// ---- Machine/FB_Centering.TcPOU
// Centraggio TL/TB di Aut260045 (ex passi 55-78 di MAIN.StateMachine, stessi numeri in nStep).
// Corsa rapida IN STROKE, ricerca dei pezzi fino a MAX STROKE con chiusura dei palpatori, arresto,
// chiusura morsa e corsa EXTRA, risalita dei centratori. Usa direttamente I/O e parametri del programma:
// e' un modulo della macchina, non del Core.
// Va chiamato a ogni ciclo PLC (gli FB di movimento e i timer devono girare sempre); con bExecute
// esegue, senza torna a Idle. Gli allarmi li memorizza qui (RaiseAlarm); il ciclo legge bDone, bFailed, bAbort.
FUNCTION_BLOCK FB_Centering
VAR_INPUT
	bExecute		: BOOL;				// il ciclo e' nel passo Centering
	bStart			: BOOL;				// consenso start (attese del passo-passo)
	bStepMode		: BOOL;				// passo-passo: tra le fasi si aspetta lo start
	fMoveSpeed		: LREAL := 200;		// velocita' USE nelle corse IN STROKE ed EXTRA
	fSearchSpeed	: LREAL := 30;		// velocita' USE nella ricerca dei pezzi
	nGroupIdBase	: UDINT := 7;		// ID NC dei gruppi da svuotare prima delle corse PTP
END_VAR
VAR_IN_OUT
	stUseL			: AXIS_REF;
	stUseR			: AXIS_REF;
END_VAR
VAR_OUTPUT
	nStep			: E_CenteringStep;
	bDone			: BOOL;		// centraggio finito: fMeasureL/R valide
	bFailed			: BOOL;		// pezzo gia' presente o non trovato: si rifa' il posizionamento iniziale
	bAbort			: BOOL;		// errore NC: il ciclo va in abort
	fMeasureL		: LREAL;	// corsa di ricerca SX (inizio - fine), per la tolleranza TB
	fMeasureR		: LREAL;
END_VAR
VAR
	fbClearGroup	: ARRAY[0..2] OF CfgReconfigGroup;
	fbMoveL			: MC_MoveAbsolute;
	fbMoveR			: MC_MoveAbsolute;
	fbStopL			: MC_Halt;
	fbStopR			: MC_Halt;
	fbClampsDelay	: TON;
	fbTlClampsDelay	: TON;
	fbUpDownDelay	: TON;
	fStrokeInL		: LREAL;
	fStrokeInR		: LREAL;
	fStartL			: LREAL;
	fStartR			: LREAL;
	fMaxStrokeL		: LREAL;
	fMaxStrokeR		: LREAL;
	fEndL			: LREAL;
	fEndR			: LREAL;
	fExtraL			: LREAL;
	fExtraR			: LREAL;
	pz1Found		: BOOL;
	pz2Found		: BOOL;
	pz3Found		: BOOL;
	pz4Found		: BOOL;
	i				: UINT;
END_VAR

// Valori di riposo a ogni ciclo (prima in MAIN.InitCyclic): i passi li riaccendono.
fbStopL.Execute := FALSE;
fbStopR.Execute := FALSE;
fbMoveL.Execute := FALSE;
fbMoveL.Velocity := 0;
fbMoveR.Execute := FALSE;
fbMoveR.Velocity := 0;
fbClampsDelay.IN := FALSE;
fbClampsDelay.PT := T#800MS;
fbTlClampsDelay.IN := FALSE;
fbTlClampsDelay.PT := T#250MS;
fbUpDownDelay.IN := FALSE;
fbUpDownDelay.PT := T#800MS;
bDone := FALSE;
bFailed := FALSE;
bAbort := FALSE;

IF NOT bExecute THEN
	nStep := E_CenteringStep.Idle;
ELSIF nStep = E_CenteringStep.Idle THEN
	nStep := E_CenteringStep.ClearGroups;
END_IF

CASE nStep OF
	(******************* Clear groups for centering *******************)  
	E_CenteringStep.ClearGroups:
		FOR i:=0 TO 2 DO
			fbClearGroup[i](
				nGroupId:=nGroupIdBase+i,
				bExecute:=TRUE,
				tTimeOut:=T#100MS );
		END_FOR
		
		IF (NOT fbClearGroup[0].bBusy) AND (NOT fbClearGroup[1].bBusy) AND (NOT fbClearGroup[2].bBusy) THEN
			fbClearGroup[0]( bExecute:=FALSE );
			fbClearGroup[1]( bExecute:=FALSE );
			fbClearGroup[2]( bExecute:=FALSE );
			nStep := E_CenteringStep.ApproachPrepare;
			
			//IO.centeringLeft1Set := FALSE;
			//IO.centeringLeft2Set := FALSE;
			//IO.centeringLeft3Set := FALSE;
			//IO.centeringLeft4Set := FALSE;
			io.centeringOutSet := TRUE;
		END_IF
		
		IF fbClearGroup[0].bErr OR fbClearGroup[1].bErr OR fbClearGroup[2].bErr THEN
			RaiseAlarm(Id := E_Alarm.NcCenteringClearGroup, Info := MAX(fbClearGroup[0].nErrId, fbClearGroup[1].nErrId, fbClearGroup[2].nErrId));
			bAbort := TRUE;
			nStep := E_CenteringStep.Error;
		END_IF
	
	(*************** Prepare fast in stroke movement ***************)  
	E_CenteringStep.ApproachPrepare:	
		fStrokeInL := stUseL.NcToPlc.ActPos - ProgramDB.parameters.inStrokeL;
		fStrokeInR := stUseR.NcToPlc.ActPos - ProgramDB.parameters.inStrokeR;
	    fbMoveL(Axis := stUseL, Execute := FALSE);
		fbMoveR(Axis := stUseR, Execute := FALSE);
		nStep := E_CenteringStep.Approach;
		
	(*************** Execute fast in stroke ***************) 
	E_CenteringStep.Approach:	
		fbMoveL.Position := fStrokeInL;
		fbMoveL.Velocity := fMoveSpeed;
		fbMoveL.Execute := TRUE;
		
		fbMoveR.Position := fStrokeInR;
		fbMoveR.Velocity := fMoveSpeed;
		fbMoveR.Execute := TRUE;
			
		IF fbMoveL.Done AND fbMoveR.Done  THEN
			IF bStart OR NOT bStepMode THEN
				nStep := E_CenteringStep.ApproachCheck;
			END_IF
		END_IF
		
		IF IO.centering1LeftIn OR IO.centering2LeftIn OR IO.centering3LeftIn THEN
			nStep := E_CenteringStep.ApproachCheck;
		END_IF
		
		IF fbMoveL.Error OR fbMoveR.Error  THEN
			RaiseAlarm(Id := E_Alarm.NcCenteringApproach, Info := MAX(fbMoveL.ErrorID, fbMoveR.ErrorID));
			bAbort := TRUE;
			nStep := E_CenteringStep.Error;
		END_IF
	
	(*************** Evaluation after in stroke ***************) 
	E_CenteringStep.ApproachCheck:	
		IF IO.centering1LeftIn OR IO.centering2LeftIn OR IO.centering3LeftIn THEN
			RaiseAlarm(Id := E_Alarm.CenteringPartAlreadyPresent, Info := 0);
			nStep := E_CenteringStep.Failed;
		ELSE
			nStep := E_CenteringStep.SearchPrepare;
		END_IF
		
	(*************** Prepare max stroke movement ***************) 
	E_CenteringStep.SearchPrepare:	
		fStartL := stUseL.NcToPlc.ActPos;
		fStartR := stUseR.NcToPlc.ActPos;
		fMaxStrokeL := fStartL - ProgramDB.parameters.maxStrokeL;
		fMaxStrokeR := fStartR - ProgramDB.parameters.maxStrokeR;
		pz1Found := FALSE;
		pz2Found := FALSE;
		pz3Found := FALSE;
		pz4Found := FALSE;
		io.centeringOutSet := FALSE;
		nStep := E_CenteringStep.Search;
		
	(*************** Execute max stroke movement ***************) 
	E_CenteringStep.Search:	
		fbMoveL.Position := fMaxStrokeL;
		fbMoveL.Velocity := fSearchSpeed;
		fbMoveL.Execute := TRUE;
		fbMoveL.Options.IgnorePositionMonitoring := TRUE;
		
		fbMoveR.Position := fMaxStrokeR;
		fbMoveR.Velocity := fSearchSpeed;
		fbMoveR.Execute := TRUE;
		fbMoveR.Options.IgnorePositionMonitoring := TRUE;
		
		IF fbMoveL.Done AND fbMoveR.Done  THEN
			RaiseAlarm(Id := E_Alarm.CenteringPartNotFound, Info := 0);
			nStep := E_CenteringStep.Failed;
		END_IF
		
		CASE ProgramDB.parameters.pcsCycle OF
			1:
				IF IO.centering1LeftIn THEN
					IO.centringClamp1Left := TRUE;
					//IO.centeringLeft1Set := TRUE;
					nStep := E_CenteringStep.StopAxes;
				END_IF
			2:
				IF IO.centering1LeftIn AND NOT pz1Found THEN
					IO.centringClamp1Left := TRUE;
					//IO.centeringLeft1Set := TRUE;
					pz1Found := TRUE;
					nStep := E_CenteringStep.PieceClamp;
				END_IF
				
				IF IO.centering2LeftIn AND NOT pz2Found THEN
					IO.centringClamp2Left := TRUE;

					//IO.centeringLeft2Set := TRUE;
					pz2Found := TRUE;
					nStep := E_CenteringStep.PieceClamp;
				END_IF
				
				IF IO.centering1LeftIn AND IO.centering2LeftIn THEN
					nStep := E_CenteringStep.StopAxes;
				END_IF
			3:
				IF IO.centering1LeftIn AND NOT pz1Found THEN
					IO.centringClamp1Left := TRUE;
					//IO.centeringLeft1Set := TRUE;
					pz1Found := TRUE;
					nStep := E_CenteringStep.PieceClamp;
				END_IF
				
				IF IO.centering2LeftIn AND NOT pz2Found THEN
					IO.centringClamp2Left := TRUE;
					//IO.centeringLeft2Set := TRUE;
					pz2Found := TRUE;
					nStep := E_CenteringStep.PieceClamp;
				END_IF
				
				IF IO.centering3LeftIn AND NOT pz3Found THEN
					IO.centringClamp3Left := TRUE;
					//IO.centeringLeft3Set := TRUE;
					pz3Found := TRUE;
					nStep := E_CenteringStep.PieceClamp;
				END_IF
				
				IF IO.centering1LeftIn AND IO.centering2LeftIn AND IO.centering3LeftIn THEN
					nStep := E_CenteringStep.StopAxes;
				END_IF
			4:
				IF IO.centering1LeftIn AND NOT pz1Found THEN
					IO.centringClamp1Left := TRUE;
					//IO.centeringLeft1Set := TRUE;
					pz1Found := TRUE;
					nStep := E_CenteringStep.PieceClamp;
				END_IF
				
				IF IO.centering2LeftIn AND NOT pz2Found THEN
					IO.centringClamp2Left := TRUE;
					//IO.centeringLeft2Set := TRUE;
					pz2Found := TRUE;
					nStep := E_CenteringStep.PieceClamp;
				END_IF
				
				IF IO.centering3LeftIn AND NOT pz3Found THEN
					IO.centringClamp3Left := TRUE;
					//IO.centeringLeft3Set := TRUE;
					pz3Found := TRUE;
					nStep := E_CenteringStep.PieceClamp;
				END_IF
				
				IF IO.centering4LeftIn AND NOT pz4Found THEN
					IO.centeringLeft4Set := TRUE;
					//IO.centringClamp4Left := TRUE;
					pz4Found := TRUE;
					nStep := E_CenteringStep.PieceClamp;
				END_IF
				
				IF IO.centering1LeftIn AND IO.centering2LeftIn AND IO.centering3LeftIn  AND IO.centering4LeftIn THEN
					nStep := E_CenteringStep.StopAxes;
				END_IF
		
		END_CASE
		IF io.centering1LeftIn THEN	
			IO.centeringLeft1Set := FALSE;
		END_IF;
		IF io.centering2LeftIn THEN	
			IO.centeringLeft2Set := FALSE;
		END_IF;
		IF io.centering3LeftIn THEN	
			IO.centeringLeft3Set := FALSE;
		END_IF;
		IF io.centering4LeftIn THEN	
			IO.centeringLeft4Set := FALSE;
		END_IF;				

		
		IF fbMoveL.Error OR fbMoveR.Error  THEN
			RaiseAlarm(Id := E_Alarm.NcCenteringSearch, Info := MAX(fbMoveL.ErrorID, fbMoveR.ErrorID));
			bAbort := TRUE;
			nStep := E_CenteringStep.Error;
		END_IF
		
	(*************** Execute max stroke movement ***************) 
	E_CenteringStep.PieceClamp:
		IO.centringClampSet := TRUE;
		fbStopL.Execute := TRUE;
		fbStopR.Execute := TRUE;
		fbTlClampsDelay.IN := TRUE;

		IF (fbStopL.Done AND fbStopR.Done)THEN
			IF fbTlClampsDelay.Q THEN
				nStep := E_CenteringStep.Search;
				io.centeringOutSet := FALSE;
			END_IF
		END_IF
				
		IF fbStopL.Error OR fbStopR.Error  THEN
			RaiseAlarm(Id := E_Alarm.NcCenteringStopSearch, Info := MAX(fbStopL.ErrorID, fbStopR.ErrorID));
			bAbort := TRUE;
			nStep := E_CenteringStep.Error;
		END_IF
		
	
	(*************** Stop execution if centering input ***************) 
	E_CenteringStep.StopAxes:
		fbStopL.Execute := TRUE;
		fbStopR.Execute := TRUE;

		IO.centringClamp1Left := FALSE;
		IO.centringClamp2Left := FALSE;
		IO.centringClamp3Left := FALSE;
		IO.centringClamp4Left := FALSE;
		
		IF (fbStopL.Done AND fbStopR.Done)THEN
			IF bStart OR NOT bStepMode THEN
				nStep := E_CenteringStep.StopDelay;
			END_IF
		END_IF
		
		IF fbStopL.Error OR fbStopR.Error  THEN
			RaiseAlarm(Id := E_Alarm.NcCenteringStop, Info := MAX(fbStopL.ErrorID, fbStopR.ErrorID));
			bAbort := TRUE;
			nStep := E_CenteringStep.Error;
		END_IF
		
	E_CenteringStep.StopDelay:
		fbTlClampsDelay.IN := TRUE;
		
		IF fbTlClampsDelay.Q THEN
			nStep := E_CenteringStep.Clamp;
		END_IF
		
	(*************** Prepare extra movement ***************)  //<--------------------- CLAMP
	E_CenteringStep.Clamp: 
		IO.centringClampSet := FALSE;
		fEndL := stUseL.NcToPlc.ActPos;
		fEndR := stUseR.NcToPlc.ActPos;
		
		fExtraL := stUseL.NcToPlc.ActPos + ProgramDB.parameters.extraL;
		fExtraR := stUseR.NcToPlc.ActPos + ProgramDB.parameters.extraR;
		
		IO.clampClosedReset := FALSE;
		IO.clampClosedSet := TRUE;
		fExtraL := stUseL.NcToPlc.ActPos + ProgramDB.parameters.extraL;

		
		fbClampsDelay.IN := TRUE;
		
		IF fbClampsDelay.Q THEN
			nStep := E_CenteringStep.Extra;
		END_IF

	(*************** Execute extra movement ***************) 
	E_CenteringStep.Extra:
		fbMoveL.Execute := TRUE;
		fbMoveL.Position := fExtraL;
		fbMoveL.Velocity := fMoveSpeed;
		
		fbMoveR.Execute := TRUE;
		fbMoveR.Position := fExtraR;
		fbMoveR.Velocity := fMoveSpeed;
		
		IF fbMoveL.Done AND fbMoveR.Done THEN
			nStep := E_CenteringStep.ResetUnits;
		END_IF
		
		IF fbMoveL.Error OR fbMoveR.Error  THEN
			RaiseAlarm(Id := E_Alarm.NcCenteringExtra, Info := MAX(fbMoveL.ErrorID, fbMoveR.ErrorID));
			bAbort := TRUE;
			nStep := E_CenteringStep.Error;
		END_IF
	
	(*************** Reset centering units ***************) 
	E_CenteringStep.ResetUnits:
		IO.centringSet := FALSE;
		IO.centringReset := TRUE;
		IO.centringClampSet := FALSE;
		IO.centringLeftUpSet := FALSE;
		IO.centringLeftUpReset := TRUE;
		IO.centringRightUpSet := FALSE;
		IO.centringRightUpReset := TRUE;
		IO.centringClamp1Left := FALSE;
		IO.centringClamp2Left := FALSE;
		IO.centringClamp3Left := FALSE;
		IO.centringClamp4Left := FALSE;
		
		fbUpDownDelay.IN := TRUE;
		
		IF fbUpDownDelay.Q THEN
			nStep := E_CenteringStep.Done;
		END_IF;

	(*************** Fine ***************)
	E_CenteringStep.Done:
		fMeasureL := fStartL - fEndL;
		fMeasureR := fStartR - fEndR;
		bDone := TRUE;

	E_CenteringStep.Failed:
		bFailed := TRUE;

	E_CenteringStep.Error:
		bAbort := TRUE;
END_CASE

// FB di movimento e timer: a ogni ciclo, dopo i passi (prima in MAIN.AxisFunctionBlocks).
fbStopL(Axis := stUseL);
fbStopR(Axis := stUseR);
fbMoveL(Axis := stUseL);
fbMoveR(Axis := stUseR);
fbClampsDelay();
fbTlClampsDelay();
fbUpDownDelay();

END_FUNCTION_BLOCK

// ---- POUs/Messages/RaiseAlarm.TcPOU
// Attiva un allarme memorizzato: resta attivo fino al Reset (ClearAlarms).
// Info = dettaglio mostrato dall'HMI (ErrorID, numero funzione M, ...); 0 = nessun dettaglio.
// Id e' un valore di E_Alarm; e' UINT perche' arriva anche dal Core (dispatcher delle funzioni M), che non conosce E_Alarm.
FUNCTION RaiseAlarm : BOOL
VAR_INPUT
	Id			: UINT;
	Info		: UDINT := 0;
END_VAR

IF Id > 0 AND Id <= Size.MAX_ALARM THEN
	IF NOT Alarms.Active[Id] THEN
		Alarms.RaisedCount := Alarms.RaisedCount + 1;
		Alarms.LastRaisedId := Id;
		Alarms.LastRaisedInfo := Info;
	END_IF
	Alarms.Active[Id] := TRUE;
	Alarms.Info[Id] := Info;
	RaiseAlarm := TRUE;
END_IF

END_FUNCTION

// ---- Core/Nc/FB_NcChannels.TcPOU
// Arresto, ripartenza e reset di tutti i canali NC insieme. Va chiamato a ogni ciclo PLC con il comando
// del ciclo; bDone e bError valgono gia' nella stessa chiamata (bBusy letto subito dopo l'esecuzione),
// cosi' il passo che lo comanda aspetta davvero la fine dell'operazione su tutti i canali.
// Con None i FB ricevono bExecute FALSE e tornano pronti per il comando successivo.
FUNCTION_BLOCK FB_NcChannels
VAR_INPUT
	eCmd			: E_NcChannelCmd;
	tTimeOut		: TIME := T#500MS;
END_VAR
VAR_IN_OUT
	aNciToPlc		: ARRAY[0..Core_Param.MAX_CHANNEL-1] OF NCTOPLC_NCICHANNEL_REF;
END_VAR
VAR_OUTPUT
	bDone			: BOOL;		// comando finito su tutti i canali, senza errori
	bError			: BOOL;		// almeno un canale in errore
	nErrorId		: UDINT;	// ErrorID piu' alto tra i canali in errore
END_VAR
VAR
	fbEStop			: ARRAY[0..Core_Param.MAX_CHANNEL-1] OF ItpEStopEx;
	fbStepOn		: ARRAY[0..Core_Param.MAX_CHANNEL-1] OF ItpStepOnAfterEStopEx;
	fbReset			: ARRAY[0..Core_Param.MAX_CHANNEL-1] OF ItpResetEx2;
	bAnyBusy		: BOOL;
	ch				: UINT;
END_VAR

bAnyBusy := FALSE;
bError := FALSE;
nErrorId := 0;

FOR ch := 0 TO Core_Param.MAX_CHANNEL - 1 DO
	fbEStop[ch](bExecute := eCmd = E_NcChannelCmd.EStop, tTimeOut := tTimeOut, sNciToPlc := aNciToPlc[ch]);
	fbStepOn[ch](bExecute := eCmd = E_NcChannelCmd.StepOn, tTimeOut := tTimeOut, sNciToPlc := aNciToPlc[ch]);
	fbReset[ch](bExecute := eCmd = E_NcChannelCmd.Reset, tTimeOut := tTimeOut, sNciToPlc := aNciToPlc[ch]);

	CASE eCmd OF
		E_NcChannelCmd.EStop:
			bAnyBusy := bAnyBusy OR fbEStop[ch].bBusy;
			IF fbEStop[ch].bErr THEN
				bError := TRUE;
				nErrorId := MAX(nErrorId, fbEStop[ch].nErrId);
			END_IF
		E_NcChannelCmd.StepOn:
			bAnyBusy := bAnyBusy OR fbStepOn[ch].bBusy;
			IF fbStepOn[ch].bErr THEN
				bError := TRUE;
				nErrorId := MAX(nErrorId, fbStepOn[ch].nErrId);
			END_IF
		E_NcChannelCmd.Reset:
			bAnyBusy := bAnyBusy OR fbReset[ch].bBusy;
			IF fbReset[ch].bErr THEN
				bError := TRUE;
				nErrorId := MAX(nErrorId, fbReset[ch].nErrId);
			END_IF
	END_CASE
END_FOR

bDone := eCmd <> E_NcChannelCmd.None AND NOT bAnyBusy AND NOT bError;

END_FUNCTION_BLOCK

// ---- Core/Axes/FB_AxisModule.TcPOU
// Un asse della macchina: potenza, reset SoE e MC, jog, calibrazione e limiti software.
// Sostituisce le cinque copie per asse di MAIN (AxisFunctionBlocks, InitCyclic, calibrazioni in Manual,
// ParameterWriteManager). Una chiamata per ciclo PLC, dopo la macchina a stati: i comandi arrivano come
// ingressi in questo ciclo, gli esiti (Done/Error) si leggono nel ciclo dopo, come prima.
// Calibrazione: MC_Home diretto alla quota, lettura dell'offset encoder, scrittura persistente,
// handshake del datum di sicurezza, impulso bCalibrated di 500 ms.
// Limiti: massimo poi minimo con MC_WriteParameter, non persistente: l'HMI li riscrive a ogni avvio e al cambio
// morsa. Con MC_WriteParameterPersistent la scrittura tornava 0x0701 su alcuni assi.
// Gli allarmi non li memorizza: li chiede con eAlarm e nAlarmInfo, la macchina sceglie il numero.
FUNCTION_BLOCK FB_AxisModule
VAR_INPUT
	// Potenza
	bPowerEnable		: BOOL;					// consenso MC_Power (motori ON, emergenza ok); l'errore dell'asse lo toglie il modulo
	fOverride			: LREAL := 100;
	bUseSoEReset		: BOOL;					// azionamento SoE reale: FB_SoEReset con potenza o reset emergenza
	bSoEResetRequest	: BOOL;					// pulsante di reset emergenza
	tPoweredOffDelay	: TIME := T#100MS;		// bPowered resta TRUE per questo tempo dopo la disabilitazione
	// Reset MC
	bResetExecute		: BOOL;
	// Jog
	bJogForward			: BOOL;
	bJogBackward		: BOOL;
	fJogVelocity		: LREAL;
	fJogAcceleration	: LREAL;
	fJogDeceleration	: LREAL;				// 0 = valore di default di MC_Jog
	fJogJerk			: LREAL;
	// Calibrazione
	bCalibrationStart	: BOOL;					// a livello: parte se il modulo e' fermo
	bUseCalibrationPos	: BOOL;					// TRUE: quota fCalibrationPos, FALSE: fHomePosition
	fCalibrationPos		: LREAL;
	fHomePosition		: LREAL;
	bDatumRequest		: BOOL;					// la sicurezza chiede il datum dopo la calibrazione
	bDatumDone			: BOOL;
	tDatumTimeOut		: TIME := T#10S;
	tReadDelay			: TIME := T#200MS;		// attesa tra homing e lettura dell'offset
	// Limiti software
	bWriteLimits		: BOOL;					// fronte: scrive fUpperLimit e fLowerLimit
	fUpperLimit			: LREAL;
	fLowerLimit			: LREAL;
	nLimitsMaxTry		: UINT := 3;			// tentativi per ogni limite prima dell'allarme
	tLimitsRetryDelay	: TIME := T#500MS;		// attesa tra un tentativo fallito e il successivo
END_VAR
VAR_IN_OUT
	stAxis				: AXIS_REF;
END_VAR
VAR_OUTPUT
	bPowered			: BOOL;					// asse abilitato (con ritardo allo spegnimento)
	bResetDone			: BOOL;
	bResetError			: BOOL;
	nResetErrorId		: UDINT;
	nCalibrationStep	: UINT;					// 0 fermo, 10 homing, 12 attesa, 15 lettura offset, 20 scrittura, 22-25 datum, 30 fine
	bCalibrated			: BOOL;					// impulso di 500 ms a calibrazione finita
	bDatumExecute		: BOOL;
	nLimitsStep			: UINT;					// 0 fermo, 10 massimo, 11 attesa, 12 minimo, 15/17 attesa nuovo tentativo
	bLimitsBusy			: BOOL;
	bLimitsError		: BOOL;					// impulso: scrittura limiti fallita
	eAlarm				: E_AxisAlarm;			// allarme chiesto in questo ciclo
	nAlarmInfo			: UDINT;
	fEncoderOffset		: LREAL;
END_VAR
VAR
	fbPower				: MC_Power;
	fbSoEReset			: FB_SoEReset;
	fbReset				: MC_Reset;
	fbJog				: MC_Jog;
	fbHome				: MC_Home;
	fbReadOffset		: MC_ReadParameter;
	fbWrite				: MC_WriteParameterPersistent;	// offset encoder della calibrazione
	fbWriteLimits		: MC_WriteParameter;			// limiti software
	fbReadDelay			: TON;
	fbDatumTimeOut		: TON;
	fbCalibratedPulse	: TP;
	fbPoweredOff		: TOF;
	fbLimitsTrigger		: R_TRIG;
	fbLimitsRetry		: TON;
	nLimitsTry			: UINT;	// tentativi falliti sul limite in scrittura
	bLimitsPending		: BOOL;	// richiesta memorizzata mentre la calibrazione e' in corso
	bCalibrationCanStart : BOOL;	// ammissione prima di acquisire eventuali nuovi limiti
END_VAR

// Valori di riposo a ogni ciclo (prima in MAIN.InitCyclic): i passi qui sotto li riaccendono.
fbHome.Execute := FALSE;
fbHome.HomingMode := MC_HomingMode.MC_Direct;
fbHome.Position := fHomePosition;
fbReadOffset.Enable := FALSE;
fbReadOffset.ReadMode := E_ReadMode.READMODE_ONCE;
fbReadOffset.ParameterNumber := MC_AxisParameter.AxisEncoderOffset;
fbWrite.Execute := FALSE;
fbWriteLimits.Execute := FALSE;
fbLimitsRetry.IN := FALSE;
fbReadDelay.IN := FALSE;
fbDatumTimeOut.IN := FALSE;
fbCalibratedPulse.IN := FALSE;
bDatumExecute := FALSE;
bLimitsError := FALSE;
eAlarm := E_AxisAlarm.None;
nAlarmInfo := 0;

//*******************************************************************************************************************
// Limiti software (prima ParameterWriteManager): massimo, attesa che il FB torni libero, minimo
//*******************************************************************************************************************
// Limiti e calibrazione non si sovrappongono: una richiesta limiti durante la calibrazione resta in attesa.
// Una calibrazione gia' ammessa in questo ciclo ha precedenza su una nuova richiesta limiti.
bCalibrationCanStart := bCalibrationStart AND nCalibrationStep = 0 AND nLimitsStep = 0
	AND NOT bLimitsPending AND NOT fbWrite.Busy AND NOT fbWrite.Done AND NOT fbWrite.Error
	AND NOT fbWriteLimits.Busy AND NOT fbWriteLimits.Done AND NOT fbWriteLimits.Error;
fbLimitsTrigger(CLK := bWriteLimits);
IF fbLimitsTrigger.Q THEN
	bLimitsPending := TRUE;
END_IF
IF bLimitsPending AND nLimitsStep = 0 AND nCalibrationStep = 0 AND NOT bCalibrationCanStart
	AND NOT fbWrite.Busy AND NOT fbWrite.Done AND NOT fbWrite.Error
	AND NOT fbWriteLimits.Busy AND NOT fbWriteLimits.Done AND NOT fbWriteLimits.Error THEN
	bLimitsPending := FALSE;
	nLimitsTry := 0;
	nLimitsStep := 10;
END_IF

// Un errore (es. 0x0701 subito dopo l'avvio) si ritenta dopo tLimitsRetryDelay; l'allarme solo all'ultimo
// tentativo, con l'ErrorID di quello.
CASE nLimitsStep OF
	10:
		fbWriteLimits.Execute := TRUE;
		fbWriteLimits.Value := fUpperLimit;
		fbWriteLimits.ParameterNumber := MC_AxisParameter.AxisMaxSoftPosLimit;
		IF fbWriteLimits.Done AND NOT fbWriteLimits.Busy THEN
			nLimitsTry := 0;
			nLimitsStep := 11;
		END_IF
		IF fbWriteLimits.Error THEN
			nLimitsTry := nLimitsTry + 1;
			IF nLimitsTry < nLimitsMaxTry THEN
				nLimitsStep := 15;
			ELSE
				nLimitsStep := 0;
				bLimitsError := TRUE;
				eAlarm := E_AxisAlarm.Limits;
				nAlarmInfo := fbWriteLimits.ErrorID;
			END_IF
		END_IF
	11:
		IF NOT fbWriteLimits.Done AND NOT fbWriteLimits.Busy THEN
			nLimitsStep := 12;
		END_IF
	12:
		fbWriteLimits.Execute := TRUE;
		fbWriteLimits.Value := fLowerLimit;
		fbWriteLimits.ParameterNumber := MC_AxisParameter.AxisMinSoftPosLimit;
		IF fbWriteLimits.Done AND NOT fbWriteLimits.Busy THEN
			nLimitsStep := 0;
		END_IF
		IF fbWriteLimits.Error THEN
			nLimitsTry := nLimitsTry + 1;
			IF nLimitsTry < nLimitsMaxTry THEN
				nLimitsStep := 17;
			ELSE
				nLimitsStep := 0;
				bLimitsError := TRUE;
				eAlarm := E_AxisAlarm.Limits;
				nAlarmInfo := fbWriteLimits.ErrorID;
			END_IF
		END_IF
	15, 17:
		// Execute resta FALSE: l'errore si azzera, poi si ripete lo stesso limite (15 -> 10, 17 -> 12).
		fbLimitsRetry.IN := TRUE;
		IF fbLimitsRetry.Q AND NOT fbWriteLimits.Error AND NOT fbWriteLimits.Busy THEN
			nLimitsStep := nLimitsStep - 5;
		END_IF
END_CASE
// Attendere anche il rilascio di Done/Error prima di ammettere un'altra scrittura.
bLimitsBusy := bLimitsPending OR nLimitsStep <> 0
	OR fbWriteLimits.Busy OR fbWriteLimits.Done OR fbWriteLimits.Error
	OR (nCalibrationStep = 0 AND (fbWrite.Busy OR fbWrite.Done OR fbWrite.Error));

//*******************************************************************************************************************
// Calibrazione (prima in MAIN.Manual, una copia per asse)
//*******************************************************************************************************************
CASE nCalibrationStep OF
	0:
		IF bCalibrationCanStart THEN
			nCalibrationStep := 10;
		END_IF
	10:
		IF bUseCalibrationPos THEN
			fbHome.Position := fCalibrationPos;
		END_IF
		fbHome.Execute := TRUE;
		IF fbHome.Done THEN
			nCalibrationStep := 12;
		END_IF
		IF fbHome.Error THEN
			nCalibrationStep := 0;
			eAlarm := E_AxisAlarm.Calibration;
			nAlarmInfo := fbHome.ErrorID;
		END_IF
	12:
		fbReadDelay.IN := TRUE;
		IF fbReadDelay.Q THEN
			nCalibrationStep := 15;
		END_IF
	15:
		fbReadOffset.Enable := TRUE;
		IF fbReadOffset.Valid THEN
			nCalibrationStep := 20;
		END_IF
		IF fbReadOffset.Error THEN
			nCalibrationStep := 0;
			eAlarm := E_AxisAlarm.Calibration;
			nAlarmInfo := fbReadOffset.ErrorID;
		END_IF
	20:
		fbWrite.Execute := TRUE;
		fbWrite.Value := fEncoderOffset;
		fbWrite.ParameterNumber := MC_AxisParameter.AxisEncoderOffset;
		IF fbWrite.Done THEN
			nCalibrationStep := 22;
		END_IF
		IF fbWrite.Error THEN
			nCalibrationStep := 0;
			eAlarm := E_AxisAlarm.Calibration;
			nAlarmInfo := fbWrite.ErrorID;
		END_IF
	22:
		IF bDatumRequest THEN
			nCalibrationStep := 25;
		ELSE
			nCalibrationStep := 30;
		END_IF
	25:
		bDatumExecute := TRUE;
		fbDatumTimeOut.IN := TRUE;
		IF bDatumDone THEN
			nCalibrationStep := 30;
		END_IF
		IF fbDatumTimeOut.Q THEN
			nCalibrationStep := 0;
			eAlarm := E_AxisAlarm.Calibration;
			nAlarmInfo := 0;
		END_IF
	30:
		fbCalibratedPulse.IN := TRUE;
		nCalibrationStep := 0;
END_CASE

//*******************************************************************************************************************
// FB dell'asse, nell'ordine di prima (AxisFunctionBlocks): jog, reset, potenza, SoE, homing, scrittura, lettura
//*******************************************************************************************************************
fbJog(
	Axis			:= stAxis,
	JogForward		:= bJogForward,
	JogBackwards	:= bJogBackward,
	Mode			:= E_JogMode.MC_JOGMODE_CONTINOUS,
	Velocity		:= fJogVelocity,
	Acceleration	:= fJogAcceleration,
	Deceleration	:= fJogDeceleration,
	Jerk			:= fJogJerk);

fbReset(Axis := stAxis, Execute := bResetExecute);
bResetDone := fbReset.Done;
bResetError := fbReset.Error;
nResetErrorId := fbReset.ErrorID;

fbPower(Axis := stAxis, Enable := bPowerEnable AND stAxis.NcToPlc.ErrorCode = 0, Enable_Positive := TRUE, Enable_Negative := TRUE, Override := fOverride);
IF bUseSoEReset THEN
	fbSoEReset(Axis := stAxis, Execute := fbPower.Enable OR bSoEResetRequest);
END_IF
fbPoweredOff(IN := NOT stAxis.Status.Disabled, PT := tPoweredOffDelay, Q => bPowered);

fbHome(Axis := stAxis);
fbWrite(Axis := stAxis);
fbWriteLimits(Axis := stAxis);
fbLimitsRetry(PT := tLimitsRetryDelay);
fbReadOffset(Axis := stAxis, Value => fEncoderOffset);
fbReadDelay(PT := tReadDelay);
fbDatumTimeOut(PT := tDatumTimeOut);
fbCalibratedPulse(PT := T#500MS, Q => bCalibrated);

END_FUNCTION_BLOCK

// ---- Core/Hmi/FB_HmiWatchdog.TcPOU
// Interfaccia viva finche' il contatore cambia almeno una volta ogni tTimeOut.
FUNCTION_BLOCK FB_HmiWatchdog
VAR_INPUT
	nCounter		: UDINT;
	tTimeOut		: TIME := T#3S;
END_VAR
VAR_OUTPUT
	bAlive			: BOOL;
END_VAR
VAR
	nLast			: UDINT;
	fbTimer			: TON;
	bSeen			: BOOL;
END_VAR

IF nCounter <> nLast THEN
	nLast := nCounter;
	bSeen := TRUE;
	fbTimer(IN := FALSE);
END_IF
fbTimer(IN := TRUE, PT := tTimeOut);
bAlive := bSeen AND NOT fbTimer.Q;

END_FUNCTION_BLOCK

// ---- Core/Hmi/FB_HmiCommandHandler.TcPOU
// Riceve i comandi dell'HMI con numero di sequenza (Hmi.Cmd): bNew vale TRUE per un ciclo quando arriva un
// comando nuovo; chi lo esegue risponde con Ack(). nAck/eResult vanno in Hmi.Sts.
// Al primo ciclo dopo l'avvio del PLC il comando presente non si esegue (si allinea nAck): niente comandi
// vecchi rieseguiti dopo un riavvio.
FUNCTION_BLOCK FB_HmiCommandHandler
VAR_INPUT
	stCmd			: ST_HmiCmd;
END_VAR
VAR_OUTPUT
	bNew			: BOOL;
	nAck			: UDINT;
	eResult			: E_HmiResult;
END_VAR
VAR
	bInit			: BOOL;
END_VAR

IF NOT bInit THEN
	bInit := TRUE;
	nAck := stCmd.nSeq;
END_IF

bNew := stCmd.nSeq <> nAck AND stCmd.eCommand <> E_HmiCommand.None;
IF stCmd.nSeq <> nAck AND stCmd.eCommand = E_HmiCommand.None THEN
	nAck := stCmd.nSeq;
	eResult := E_HmiResult.UnknownCommand;
END_IF

// Risposta al comando nuovo di questo ciclo.
METHOD Ack
VAR_INPUT
	eAnswer		: E_HmiResult;
END_VAR
nAck := stCmd.nSeq;
eResult := eAnswer;
bNew := FALSE;
END_METHOD

END_FUNCTION_BLOCK

// ---- Machine/FB_MachineConfig.TcPOU
// Configurazione di Aut260045 per il Core: valvole (uscite e conferme) e tabella delle funzioni M.
// E' il solo punto da toccare per una valvola o una funzione M nuova. Si chiama a ogni ciclo, prima
// del dispatcher: i puntatori seguono gli spostamenti di memoria di un online change e la tabella
// e' sempre quella scritta qui.
// Tempi, conferme e allarmi sono quelli del vecchio MacroManager (tabella di confronto in
// _verifica_plc\macrotable). Le conferme "uguali all'uscita" sono le valvole senza sensore.
FUNCTION_BLOCK FB_MachineConfig
VAR
	stDef			: ST_MFuncDef;
END_VAR

//*******************************************************************************************************************
// Assi dei programmi (AXIS_ENUM): nome, scala velocita' (fVelo = speed * scala), correzione centraggio TB,
// quota sempre 0 (asse simulato), asse NC. Un asse nuovo (es. trascinamento): valore in AXIS_ENUM, asse NC, una riga qui.
//*******************************************************************************************************************
Axis(AXIS_ENUM.USEL,	'USE SX',		10.0,	TRUE,	FALSE,	MAIN.USEL);
Axis(AXIS_ENUM.USER,	'USE DX',		10.0,	TRUE,	FALSE,	MAIN.USER);
Axis(AXIS_ENUM.ERL,		'ER SX',		10.8,	FALSE,	FALSE,	MAIN.ERL);
Axis(AXIS_ENUM.ERR,		'ER DX',		10.8,	FALSE,	FALSE,	MAIN.ERR);
Axis(AXIS_ENUM.UR2,		'UR2',			10.8,	FALSE,	FALSE,	MAIN.UR2);
Axis(AXIS_ENUM.UR_SIM,	'UR simulato',	10.8,	FALSE,	TRUE,	MAIN.UR_SIM);

// Movimento manuale e servizio: selettore volantino, jog (velocita', accelerazione, decelerazione, jerk),
// azionamento SoE, allarmi di calibrazione e di scrittura limiti. Valori di prima (InitCyclic, Manual).
AxisService(AXIS_ENUM.ERL,		1,	100,	500,	0,		20000,	TRUE,	E_Alarm.HomingErl,	E_Alarm.ParamWriteErl);
AxisService(AXIS_ENUM.USEL,		2,	250,	500,	500,	5000,	TRUE,	E_Alarm.HomingUsel,	E_Alarm.ParamWriteUsel);
AxisService(AXIS_ENUM.UR2,		3,	100,	500,	0,		5000,	TRUE,	E_Alarm.HomingUr2,	E_Alarm.ParamWriteUr2);
AxisService(AXIS_ENUM.UR_SIM,	3,	100,	500,	0,		5000,	FALSE,	0,					0);
AxisService(AXIS_ENUM.ERR,		4,	100,	500,	0,		20000,	TRUE,	E_Alarm.HomingErr,	E_Alarm.ParamWriteErr);
AxisService(AXIS_ENUM.USER,		5,	250,	500,	0,		5000,	TRUE,	E_Alarm.HomingUser,	E_Alarm.ParamWriteUser);

// Pulsanti del volantino: per ogni posizione del selettore, la valvola del pulsante 1 e quella del pulsante 3.
Mach.aMpgButton[1, 1] := E_Valve.ErLeft;			Mach.aMpgButton[1, 2] := E_Valve.UseLeftUp;
Mach.aMpgButton[2, 1] := E_Valve.CenteringLeftUp;	Mach.aMpgButton[2, 2] := E_Valve.SupportLeft;
Mach.aMpgButton[3, 1] := E_Valve.Eject;				Mach.aMpgButton[3, 2] := E_Valve.Clamp;
Mach.aMpgButton[4, 1] := E_Valve.ErRight;			Mach.aMpgButton[4, 2] := E_Valve.UseRightUp;
Mach.aMpgButton[5, 1] := E_Valve.CenteringRightUp;	Mach.aMpgButton[5, 2] := E_Valve.SupportRight;

//*******************************************************************************************************************
// Valvole: uscita set, uscita reset (0 = monostabile), conferma set, conferma reset
//*******************************************************************************************************************
Valve(E_Valve.ErLeft,		'ER SX testa',			OUTPUT_ENUM.BISTABLE,	ADR(IO.erLeftOutSet),		ADR(IO.erLeftOutReset),		ADR(IO.erLeftOut),			ADR(IO.erLeftIn));
Valve(E_Valve.UseLeftUp,	'ER SX trasversale',	OUTPUT_ENUM.BISTABLE,	ADR(IO.useLeftUpSet),		ADR(IO.useLeftUpReset),		ADR(IO.useLeftUp),			ADR(IO.useLeftDown));
Valve(E_Valve.SupportLeft,	'Spallamento SX',		OUTPUT_ENUM.BISTABLE,	ADR(IO.supportLeftOutSet),	ADR(IO.supportLeftOutReset),	ADR(IO.supportLeftOutSet),	ADR(IO.supportLeftOutReset));
Valve(E_Valve.EpLeftBend,	'EP SX trazione',		OUTPUT_ENUM.MONOSTABLE,	ADR(IO.epLeftBend),			0,							ADR(IO.epLeftBendDown),		ADR(IO.epLeftBendUp));
Valve(E_Valve.EpLeftOut,	'EP SX estrazione',		OUTPUT_ENUM.BISTABLE,	ADR(IO.epLeftOutSet),		ADR(IO.epLeftOutReset),		ADR(IO.epLeftOut),			ADR(IO.epLeftIn));
Valve(E_Valve.ErRight,		'ER DX testa',			OUTPUT_ENUM.BISTABLE,	ADR(IO.erRightOutSet),		ADR(IO.erRightOutReset),	ADR(IO.erRightOut),			ADR(IO.erRightIn));
Valve(E_Valve.UseRightUp,	'ER DX trasversale',	OUTPUT_ENUM.BISTABLE,	ADR(IO.useRightUpSet),		ADR(IO.useRightUpReset),	ADR(IO.useRighttUp),		ADR(IO.useRightDown));
Valve(E_Valve.SupportRight,	'Spallamento DX',		OUTPUT_ENUM.BISTABLE,	ADR(IO.supportRightOutSet),	ADR(IO.supportRightOutReset),	ADR(IO.supportRightOutSet),	ADR(IO.supportRightOutReset));
Valve(E_Valve.EpRightBend,	'EP DX trazione',		OUTPUT_ENUM.MONOSTABLE,	ADR(IO.epRightBend),		0,							ADR(IO.epRightBendDown),	ADR(IO.epRightBendUp));
Valve(E_Valve.EpRightOut,	'EP DX estrazione',		OUTPUT_ENUM.BISTABLE,	ADR(IO.epRightOutSet),		ADR(IO.epRightOutReset),	ADR(IO.epRightOut),			ADR(IO.epRightIn));
Valve(E_Valve.Clamp,		'Morsa',				OUTPUT_ENUM.BISTABLE,	ADR(IO.clampClosedSet),		ADR(IO.clampClosedReset),	ADR(IO.clampClosedSet),		ADR(IO.clampClosedReset));
Valve(E_Valve.Eject,		'Espulsore',			OUTPUT_ENUM.BISTABLE,	ADR(IO.clampEjectSet),		ADR(IO.clampEjectReset),	ADR(IO.clampEjectSet),		ADR(IO.clampEjectReset));
Valve(E_Valve.CenteringLeftUp,	'Centratore SX su',	OUTPUT_ENUM.BISTABLE,	ADR(IO.centringLeftUpSet),	ADR(IO.centringLeftUpReset),	ADR(IO.centringLeftUpSet),	ADR(IO.centringLeftUpReset));
Valve(E_Valve.CenteringRightUp,	'Centratore DX su',	OUTPUT_ENUM.BISTABLE,	ADR(IO.centringRightUpSet),	ADR(IO.centringRightUpReset),	ADR(IO.centringRightUpSet),	ADR(IO.centringRightUpReset));
Valve(E_Valve.CenteringUp,		'Centratori su',		OUTPUT_ENUM.BISTABLE,	ADR(IO.centringSet),		ADR(IO.centringReset),		ADR(IO.centringSet),		ADR(IO.centringReset));
Valve(E_Valve.CenteringClamp,	'Bloccaggio centratori',	OUTPUT_ENUM.MONOSTABLE,	ADR(IO.centringClampSet),	0,						ADR(IO.centringClampSet),	ADR(IO.centringClampSet));
Valve(E_Valve.CenteringOut,		'Supporto centraggio',	OUTPUT_ENUM.MONOSTABLE,	ADR(IO.centeringOutSet),	0,							ADR(IO.centeringOutSet),	ADR(IO.centeringOutSet));
Valve(E_Valve.CenteringPiece1,	'Palpatore 1',			OUTPUT_ENUM.MONOSTABLE,	ADR(IO.centringClamp1Left),	0,							ADR(IO.centringClamp1Left),	ADR(IO.centringClamp1Left));
Valve(E_Valve.CenteringPiece2,	'Palpatore 2',			OUTPUT_ENUM.MONOSTABLE,	ADR(IO.centringClamp2Left),	0,							ADR(IO.centringClamp2Left),	ADR(IO.centringClamp2Left));
Valve(E_Valve.CenteringPiece3,	'Palpatore 3',			OUTPUT_ENUM.MONOSTABLE,	ADR(IO.centringClamp3Left),	0,							ADR(IO.centringClamp3Left),	ADR(IO.centringClamp3Left));
Valve(E_Valve.CenteringPiece4,	'Palpatore 4',			OUTPUT_ENUM.MONOSTABLE,	ADR(IO.centringClamp4Left),	0,							ADR(IO.centringClamp4Left),	ADR(IO.centringClamp4Left));
Valve(E_Valve.CenteringAir1,	'Esclusione aria 1',	OUTPUT_ENUM.MONOSTABLE,	ADR(IO.centeringLeft1Set),	0,							ADR(IO.centeringLeft1Set),	ADR(IO.centeringLeft1Set));
Valve(E_Valve.CenteringAir2,	'Esclusione aria 2',	OUTPUT_ENUM.MONOSTABLE,	ADR(IO.centeringLeft2Set),	0,							ADR(IO.centeringLeft2Set),	ADR(IO.centeringLeft2Set));
Valve(E_Valve.CenteringAir3,	'Esclusione aria 3',	OUTPUT_ENUM.MONOSTABLE,	ADR(IO.centeringLeft3Set),	0,							ADR(IO.centeringLeft3Set),	ADR(IO.centeringLeft3Set));
Valve(E_Valve.CenteringAir4,	'Esclusione aria 4',	OUTPUT_ENUM.MONOSTABLE,	ADR(IO.centeringLeft4Set),	0,							ADR(IO.centeringLeft4Set),	ADR(IO.centeringLeft4Set));

//*******************************************************************************************************************
// Ingressi mostrati all'HMI (sensori)
//*******************************************************************************************************************
Input(1,	'ER SX dentro',			ADR(IO.erLeftIn));
Input(2,	'ER SX fuori',			ADR(IO.erLeftOut));
Input(3,	'ER SX trasv. su',		ADR(IO.useLeftUp));
Input(4,	'ER SX trasv. giu',		ADR(IO.useLeftDown));
Input(5,	'ER DX dentro',			ADR(IO.erRightIn));
Input(6,	'ER DX fuori',			ADR(IO.erRightOut));
Input(7,	'ER DX trasv. su',		ADR(IO.useRighttUp));
Input(8,	'ER DX trasv. giu',		ADR(IO.useRightDown));
Input(9,	'Centratore pezzo 1',	ADR(IO.centering1LeftIn));
Input(10,	'Centratore pezzo 2',	ADR(IO.centering2LeftIn));
Input(11,	'Centratore pezzo 3',	ADR(IO.centering3LeftIn));
Input(12,	'Centratore pezzo 4',	ADR(IO.centering4LeftIn));
Input(13,	'EP SX dentro',			ADR(IO.epLeftIn));
Input(14,	'EP SX fuori',			ADR(IO.epLeftOut));
Input(15,	'EP SX trazione giu',	ADR(IO.epLeftBendDown));
Input(16,	'EP SX trazione su',	ADR(IO.epLeftBendUp));
Input(17,	'EP DX dentro',			ADR(IO.epRightIn));
Input(18,	'EP DX fuori',			ADR(IO.epRightOut));
Input(19,	'EP DX trazione giu',	ADR(IO.epRightBendDown));
Input(20,	'EP DX trazione su',	ADR(IO.epRightBendUp));

//*******************************************************************************************************************
// Funzioni M. Canali: 0 = unita' SX, 1 = unita' DX, 2 = UR2.
//*******************************************************************************************************************
Mach.nMFuncCount := 0;

// --- Canale 0, unita' SX ---
AddMFunc(F_MSync(0, 62, 0, 0, Mach.SYNC_ACK_L, 0, 0, 0, 0));													// USE SX in posizione
AddMFunc(F_MSync(0, 61, Mach.SYNC_ACK_R, 0, 0, Mach.SYNC_ACK_R, 0, 0, E_Alarm.SyncLeftWaitRight));			// aspetta la USE DX
AddMFunc(F_MSync(0, 80, Mach.SYNC_UR2_DONE, 0, 0, 0, 0, Mach.SYNC_UR2_ACK_L, E_Alarm.SyncLeftWaitUr2));		// aspetta l'UR2
AddMFunc(F_MSync(0, 112, 0, Mach.SYNC_UR2_DONE, 0, Mach.SYNC_UR2_ACK_L, Mach.SYNC_UR2_ACK_L, 0, E_Alarm.SyncLeftWaitUr2Ack));	// conferma all'UR2
AddMFunc(F_MSync(0, 150, 0, 0, 0, Mach.SYNC_UR2_ACK_L OR Mach.SYNC_DONE_L, 0, 0, 0));							// reset sincronismi
AddMFunc(F_MValve(0, 40, E_Valve.ErLeft,		OUTPUT_ACTION_ENUM.SET,		T#1000MS, T#500MS,	E_Alarm.ErLeftUp));
AddMFunc(F_MValve(0, 41, E_Valve.ErLeft,		OUTPUT_ACTION_ENUM.RESET,	T#2000MS, T#500MS,	E_Alarm.ErLeftDown));
AddMFunc(F_MValve(0, 44, E_Valve.UseLeftUp,	OUTPUT_ACTION_ENUM.SET,		T#3000MS, T#500MS,	E_Alarm.UseLeftUp));
AddMFunc(F_MValve(0, 45, E_Valve.UseLeftUp,	OUTPUT_ACTION_ENUM.RESET,	T#2000MS, T#230MS,	E_Alarm.UseLeftDown));
AddMFunc(F_MValveDirect(0, 54, E_Valve.UseLeftUp, OUTPUT_ACTION_ENUM.SET));
AddMFunc(F_MValveDirect(0, 55, E_Valve.UseLeftUp, OUTPUT_ACTION_ENUM.RESET));
AddMFunc(F_MValve(0, 50, E_Valve.SupportLeft,	OUTPUT_ACTION_ENUM.SET,		T#2000MS, T#400MS,	E_Alarm.SupportLeftOut));
AddMFunc(F_MValve(0, 51, E_Valve.SupportLeft,	OUTPUT_ACTION_ENUM.RESET,	T#2000MS, T#400MS,	E_Alarm.SupportLeftIn));
AddMFunc(F_MValve(0, 70, E_Valve.EpLeftBend,	OUTPUT_ACTION_ENUM.SET,		T#2000MS, T#100MS,	E_Alarm.EpLeftBend));
AddMFunc(F_MValve(0, 72, E_Valve.EpLeftOut,	OUTPUT_ACTION_ENUM.SET,		T#2000MS, T#100MS,	E_Alarm.EpLeftOut));
AddMFunc(F_MValve(0, 73, E_Valve.EpLeftOut,	OUTPUT_ACTION_ENUM.RESET,	T#2000MS, T#100MS,	E_Alarm.EpLeftIn));
AddMFunc(F_MValve(0, 74, E_Valve.EpLeftBend,	OUTPUT_ACTION_ENUM.RESET,	T#2000MS, T#1000MS,	E_Alarm.EpLeftBendReturn));
AddMFunc(F_MSimple(0, 95, E_MFuncKind.WaitStart));
AddMFunc(F_MSimple(0, 130, E_MFuncKind.WaitH));
AddMFunc(F_MSimple(0, 135, E_MFuncKind.LineNo));
AddMFunc(F_MSimple(0, 140, E_MFuncKind.Nop));

// --- Canale 1, unita' DX ---
AddMFunc(F_MSync(1, 63, 0, 0, Mach.SYNC_ACK_R, 0, 0, 0, 0));													// USE DX in posizione
AddMFunc(F_MSync(1, 60, Mach.SYNC_ACK_L, 0, 0, Mach.SYNC_ACK_L, 0, 0, E_Alarm.SyncRightWaitLeft));			// aspetta la USE SX
AddMFunc(F_MSync(1, 80, Mach.SYNC_UR2_DONE, 0, 0, 0, 0, Mach.SYNC_UR2_ACK_R, E_Alarm.SyncRightWaitUr2));		// aspetta l'UR2
AddMFunc(F_MSync(1, 113, 0, Mach.SYNC_UR2_DONE, 0, Mach.SYNC_UR2_ACK_R, Mach.SYNC_UR2_ACK_R, 0, E_Alarm.SyncRightWaitUr2Ack));	// conferma all'UR2
AddMFunc(F_MSync(1, 150, 0, 0, 0, Mach.SYNC_UR2_ACK_R OR Mach.SYNC_DONE_R, 0, 0, 0));							// reset sincronismi
AddMFunc(F_MValve(1, 42, E_Valve.ErRight,		OUTPUT_ACTION_ENUM.SET,		T#1000MS, T#300MS,	E_Alarm.ErRightUp));
AddMFunc(F_MValve(1, 43, E_Valve.ErRight,		OUTPUT_ACTION_ENUM.RESET,	T#1000MS, T#100MS,	E_Alarm.ErRightDown));
AddMFunc(F_MValve(1, 46, E_Valve.UseRightUp,	OUTPUT_ACTION_ENUM.SET,		T#2000MS, T#400MS,	E_Alarm.UseRightUp));
AddMFunc(F_MValve(1, 47, E_Valve.UseRightUp,	OUTPUT_ACTION_ENUM.RESET,	T#2000MS, T#400MS,	E_Alarm.UseRightDown));
AddMFunc(F_MValveDirect(1, 56, E_Valve.UseRightUp, OUTPUT_ACTION_ENUM.SET));
AddMFunc(F_MValveDirect(1, 57, E_Valve.UseRightUp, OUTPUT_ACTION_ENUM.RESET));
AddMFunc(F_MValve(1, 48, E_Valve.SupportRight,	OUTPUT_ACTION_ENUM.SET,		T#2000MS, T#200MS,	E_Alarm.SupportRightOut));
AddMFunc(F_MValve(1, 49, E_Valve.SupportRight,	OUTPUT_ACTION_ENUM.RESET,	T#2000MS, T#100MS,	E_Alarm.SupportRightIn));
AddMFunc(F_MValve(1, 70, E_Valve.EpRightBend,	OUTPUT_ACTION_ENUM.SET,		T#2000MS, T#100MS,	E_Alarm.EpRightBend));
AddMFunc(F_MValve(1, 72, E_Valve.EpRightOut,	OUTPUT_ACTION_ENUM.SET,		T#2000MS, T#100MS,	E_Alarm.EpRightOut));
AddMFunc(F_MValve(1, 73, E_Valve.EpRightOut,	OUTPUT_ACTION_ENUM.RESET,	T#2000MS, T#100MS,	E_Alarm.EpRightIn));
AddMFunc(F_MValve(1, 74, E_Valve.EpRightBend,	OUTPUT_ACTION_ENUM.RESET,	T#2000MS, T#1000MS,	E_Alarm.EpRightBendReturn));
AddMFunc(F_MSimple(1, 96, E_MFuncKind.WaitStart));
AddMFunc(F_MSimple(1, 130, E_MFuncKind.WaitH));
AddMFunc(F_MSimple(1, 135, E_MFuncKind.LineNo));
AddMFunc(F_MSimple(1, 140, E_MFuncKind.Nop));

// --- Canale 2, UR2 ---
AddMFunc(F_MSync(2, 78, 0, 0, Mach.SYNC_UR2_DONE, 0, 0, 0, 0));													// UR2 in posizione
AddMFunc(F_MSync(2, 110, Mach.SYNC_UR2_ACK_L OR Mach.SYNC_UR2_ACK_R, 0, 0, Mach.SYNC_UR2_DONE, 0, 0, E_Alarm.SyncUr2WaitUseAck));	// aspetta la conferma delle USE
AddMFunc(F_MSync(2, 116, Mach.SYNC_ACK_L OR Mach.SYNC_ACK_R, 0, 0, Mach.SYNC_ACK_L OR Mach.SYNC_ACK_R, 0, 0, E_Alarm.SyncUr2WaitUse));	// aspetta le due USE
AddMFunc(F_MSync(2, 150, 0, 0, 0, Mach.SYNC_ACK_UR2 OR Mach.SYNC_UR2_DONE OR Mach.SYNC_UR2_REQ_L OR Mach.SYNC_UR2_REQ_R, 0, 0, 0));	// reset sincronismi

// Morsa: la conferma e' l'uscita stessa, il timeout non puo' scattare (Ignore come prima).
stDef := F_MValve(2, 100, E_Valve.Clamp,	OUTPUT_ACTION_ENUM.SET,		T#1000MS, T#300MS,	0);
stDef.eOnError := E_MFuncOnError.Ignore;
AddMFunc(stDef);
stDef := F_MValve(2, 101, E_Valve.Clamp,	OUTPUT_ACTION_ENUM.RESET,	T#500MS, T#500MS,	0);
stDef.eOnError := E_MFuncOnError.Ignore;
AddMFunc(stDef);

// Espulsione: parte solo con l'UR2 a zero (altrimenti attesa con time-out, allarme 128);
// se l'espulsore non conferma la funzione viene concessa lo stesso, senza allarme (come prima).
stDef := F_MValve(2, 102, E_Valve.Eject,	OUTPUT_ACTION_ENUM.SET,		T#500MS, T#500MS,	0);
stDef.eOnError := E_MFuncOnError.Grant;
stDef.nInterlock := Mach.IL_UR2_AT_ZERO;
stDef.nWaitAlarmId := E_Alarm.EjectUr2NotAtZero;
AddMFunc(stDef);

// Ritorno espulsore: il post-delay e' il parametro H della riga (DeltaT di espulsione).
stDef := F_MValve(2, 103, E_Valve.Eject,	OUTPUT_ACTION_ENUM.RESET,	T#1000MS, T#0MS,	0);
stDef.bPostDelayFromH := TRUE;
stDef.eOnError := E_MFuncOnError.Ignore;
AddMFunc(stDef);

AddMFunc(F_MSimple(2, 97, E_MFuncKind.WaitStart));
AddMFunc(F_MSimple(2, 130, E_MFuncKind.WaitH));
AddMFunc(F_MSimple(2, 135, E_MFuncKind.LineNo));
AddMFunc(F_MSimple(2, 140, E_MFuncKind.Nop));

// Aggiunge una riga alla tabella delle funzioni M (oltre MAX_MFUNC la riga si perde: aumentare Mach.MAX_MFUNC).
METHOD PRIVATE AddMFunc
VAR_INPUT
	stNew		: ST_MFuncDef;
END_VAR
IF Mach.nMFuncCount < Mach.MAX_MFUNC THEN
	Mach.nMFuncCount := Mach.nMFuncCount + 1;
	Mach.aMFunc[Mach.nMFuncCount] := stNew;
END_IF
END_METHOD

// Descrive un asse dei programmi e ne copia ID NC e posizione attuale (a ogni ciclo).
METHOD PRIVATE Axis
VAR_INPUT
	eAxis					: AXIS_ENUM;
	sName					: STRING(23);
	fSpeedScale				: LREAL;
	bCenteringCorrection	: BOOL;
	bTargetZero				: BOOL;
END_VAR
VAR_IN_OUT
	stAxis					: AXIS_REF;
END_VAR
VAR
	n						: UINT;
END_VAR
n := TO_UINT(eAxis);
Mach.aAxisCfg[n].bDefined := TRUE;
Mach.aAxisCfg[n].sName := sName;
Mach.aAxisCfg[n].fSpeedScale := fSpeedScale;
Mach.aAxisCfg[n].bCenteringCorrection := bCenteringCorrection;
Mach.aAxisCfg[n].bTargetZero := bTargetZero;
Mach.aAxisCfg[n].nNcAxisId := stAxis.NcToPlc.AxisId;
Mach.aAxisCfg[n].fActPos := stAxis.NcToPlc.ActPos;
Mach.aAxisCfg[n].fActVelo := stAxis.NcToPlc.ActVelo;
Mach.aAxisCfg[n].nErrorCode := stAxis.NcToPlc.ErrorCode;
Mach.aAxisCfg[n].bDisabled := stAxis.Status.Disabled;
Mach.aAxisCfg[n].bMoving := stAxis.Status.Moving;
END_METHOD

// Movimento manuale e servizio di un asse (FB_AxisModule).
METHOD PRIVATE AxisService
VAR_INPUT
	eAxis				: AXIS_ENUM;
	nMpgSelector		: UINT;
	fJogVelocity		: LREAL;
	fJogAcceleration	: LREAL;
	fJogDeceleration	: LREAL;
	fJogJerk			: LREAL;
	bSoEReset			: BOOL;
	nCalibrationAlarmId	: UINT;
	nLimitsAlarmId		: UINT;
END_VAR
VAR
	n					: UINT;
END_VAR
n := TO_UINT(eAxis);
Mach.aAxisCfg[n].nMpgSelector := nMpgSelector;
Mach.aAxisCfg[n].fJogVelocity := fJogVelocity;
Mach.aAxisCfg[n].fJogAcceleration := fJogAcceleration;
Mach.aAxisCfg[n].fJogDeceleration := fJogDeceleration;
Mach.aAxisCfg[n].fJogJerk := fJogJerk;
Mach.aAxisCfg[n].bSoEReset := bSoEReset;
Mach.aAxisCfg[n].nCalibrationAlarmId := nCalibrationAlarmId;
Mach.aAxisCfg[n].nLimitsAlarmId := nLimitsAlarmId;
END_METHOD

// Descrive un ingresso mostrato all'HMI.
METHOD PRIVATE Input
VAR_INPUT
	nIndex		: UINT;
	sName		: STRING(23);
	pInput		: POINTER TO BOOL;
END_VAR
Mach.aInput[nIndex].sName := sName;
Mach.aInput[nIndex].pInput := pInput;
END_METHOD

// Descrive una valvola: uscite e conferme (pReset = 0 per la monostabile).
METHOD PRIVATE Valve
VAR_INPUT
	eValve		: E_Valve;
	sName		: STRING(23);
	eType		: OUTPUT_ENUM;
	pSet		: POINTER TO BOOL;
	pReset		: POINTER TO BOOL;
	pFbSet		: POINTER TO BOOL;
	pFbReset	: POINTER TO BOOL;
END_VAR
Mach.aValve[eValve].sName := sName;
Mach.aValve[eValve].eType := eType;
Mach.aValve[eValve].pSet := pSet;
Mach.aValve[eValve].pReset := pReset;
Mach.aValve[eValve].pFbSet := pFbSet;
Mach.aValve[eValve].pFbReset := pFbReset;
END_METHOD

END_FUNCTION_BLOCK

// ---- Core/Sync/F_MSync.TcPOU
// Funzione M di sincronismo tra canali sui bit di un DWORD comune.
// A ogni ciclo in cui e' richiesta: dwSetWhileWaiting a 1, dwClearWhileWaiting a 0.
// Concessa quando i bit di dwWaitSet sono tutti a 1 e quelli di dwWaitClear tutti a 0;
// alla concessione dwSetOnGrant a 1 e dwClearOnGrant a 0.
FUNCTION F_MSync : ST_MFuncDef
VAR_INPUT
	nChannel			: UINT;
	nMFunc				: UINT;
	dwWaitSet			: DWORD;
	dwWaitClear			: DWORD;
	dwSetOnGrant		: DWORD;
	dwClearOnGrant		: DWORD;
	dwSetWhileWaiting	: DWORD;
	dwClearWhileWaiting	: DWORD;
	nWaitAlarmId		: UINT;		// allarme di time-out dell'attesa, 0 = nessuno
END_VAR

F_MSync.nChannel := nChannel;
F_MSync.nMFunc := nMFunc;
F_MSync.eKind := E_MFuncKind.Sync;
F_MSync.dwWaitSet := dwWaitSet;
F_MSync.dwWaitClear := dwWaitClear;
F_MSync.dwSetOnGrant := dwSetOnGrant;
F_MSync.dwClearOnGrant := dwClearOnGrant;
F_MSync.dwSetWhileWaiting := dwSetWhileWaiting;
F_MSync.dwClearWhileWaiting := dwClearWhileWaiting;
F_MSync.nWaitAlarmId := nWaitAlarmId;

END_FUNCTION

// ---- Core/Sync/F_MValve.TcPOU
// Funzione M che muove una valvola e aspetta la conferma; in caso di timeout allarme e abort.
FUNCTION F_MValve : ST_MFuncDef
VAR_INPUT
	nChannel	: UINT;
	nMFunc		: UINT;
	nValve		: UINT;
	eAction		: OUTPUT_ACTION_ENUM;
	tTimeout	: TIME;
	tPostDelay	: TIME;
	nAlarmId	: UINT;
END_VAR

F_MValve.nChannel := nChannel;
F_MValve.nMFunc := nMFunc;
F_MValve.eKind := E_MFuncKind.Valve;
F_MValve.nValve := nValve;
F_MValve.eAction := eAction;
F_MValve.tTimeout := tTimeout;
F_MValve.tPostDelay := tPostDelay;
F_MValve.nAlarmId := nAlarmId;
F_MValve.eOnError := E_MFuncOnError.Abort;

END_FUNCTION

// ---- Core/Sync/F_MValveDirect.TcPOU
// Funzione M che scrive le uscite di una valvola e viene concessa subito, senza aspettare la conferma.
FUNCTION F_MValveDirect : ST_MFuncDef
VAR_INPUT
	nChannel	: UINT;
	nMFunc		: UINT;
	nValve		: UINT;
	eAction		: OUTPUT_ACTION_ENUM;
END_VAR

F_MValveDirect.nChannel := nChannel;
F_MValveDirect.nMFunc := nMFunc;
F_MValveDirect.eKind := E_MFuncKind.ValveDirect;
F_MValveDirect.nValve := nValve;
F_MValveDirect.eAction := eAction;

END_FUNCTION

// ---- Core/Sync/F_MSimple.TcPOU
// Funzione M senza parametri: Nop, WaitH, LineNo, WaitStart.
FUNCTION F_MSimple : ST_MFuncDef
VAR_INPUT
	nChannel	: UINT;
	nMFunc		: UINT;
	eKind		: E_MFuncKind;
END_VAR

F_MSimple.nChannel := nChannel;
F_MSimple.nMFunc := nMFunc;
F_MSimple.eKind := eKind;

END_FUNCTION

// ---- Core/Sync/FB_MFuncDispatcher.TcPOU
// Esegue le funzioni M con handshake chieste dai canali NC, secondo la tabella aDef della macchina.
// Una chiamata per ciclo PLC. Per ogni canale: se c'e' una richiesta (e non e' appena stata concessa)
// cerca la riga (canale, M) e la esegue; senza riga chiede l'allarme nUnknownAlarmId (Info = canale*1000 + M,
// canale contato da 1) e l'abort. Non scrive allarmi ne' passi del ciclo: li chiede con bAbort e aAlarmId,
// la macchina decide (MAIN.MacroManager).
// Dopo la concessione il canale resta escluso per 10 ms, il tempo che l'NC abbassi la richiesta.
FUNCTION_BLOCK FB_MFuncDispatcher
VAR_INPUT
	bStart				: BOOL;		// consenso start per le funzioni WaitStart (passo-passo)
	bCycleRunning		: BOOL;		// ciclo in corso: solo allora una M sconosciuta chiede l'abort
	nUnknownAlarmId		: UINT;		// allarme per una M senza riga in tabella
	nDefCount			: UINT;		// righe valide di aDef, a partire dal primo indice
END_VAR
VAR_IN_OUT
	aNciToPlc			: ARRAY[0..Core_Param.MAX_CHANNEL-1] OF NCTOPLC_NCICHANNEL_REF;
	aPlcToNci			: ARRAY[0..Core_Param.MAX_CHANNEL-1] OF PLCTONC_NCICHANNEL_REF;
	aDef				: ARRAY[*] OF ST_MFuncDef;
	aValve				: ARRAY[*] OF ST_Valve;
	aInterlock			: ARRAY[*] OF BOOL;
	dwSyncFlags			: DWORD;
END_VAR
VAR_OUTPUT
	bAbort				: BOOL;		// in questo ciclo una funzione M chiede l'abort del ciclo
	aAlarmId			: ARRAY[0..Core_Param.MAX_CHANNEL-1] OF UINT;		// allarme da memorizzare, 0 = nessuno
	aAlarmInfo			: ARRAY[0..Core_Param.MAX_CHANNEL-1] OF UDINT;
	aWaiting			: ARRAY[0..Core_Param.MAX_CHANNEL-1] OF BOOL;		// fermo su un'attesa con time-out (sync o interlock)
	aWaitAlarmId		: ARRAY[0..Core_Param.MAX_CHANNEL-1] OF UINT;		// allarme di quell'attesa
	aLineNo				: ARRAY[0..Core_Param.MAX_CHANNEL-1] OF UDINT;	// ultima riga del programma (funzione LineNo)
END_VAR
VAR
	fbSetMacro			: ARRAY[0..Core_Param.MAX_CHANNEL-1] OF SetMacro;
	fbWaitMacro			: ARRAY[0..Core_Param.MAX_CHANNEL-1] OF WaitMacro;
	fbGrantTrig			: ARRAY[0..Core_Param.MAX_CHANNEL-1] OF R_TRIG;
	fbGrantHold			: ARRAY[0..Core_Param.MAX_CHANNEL-1] OF TOF;
	aNoResetOutput		: ARRAY[0..Core_Param.MAX_CHANNEL-1] OF BOOL;	// uscita "reset" fittizia per le valvole monostabili
	ch					: UINT;
	i					: DINT;
	nDef				: DINT;
	nMFunc				: UINT;
	bGrant				: BOOL;
	stDef				: ST_MFuncDef;
	stValve				: ST_Valve;
END_VAR

bAbort := FALSE;

FOR ch := 0 TO Core_Param.MAX_CHANNEL - 1 DO
	aAlarmId[ch] := 0;
	aAlarmInfo[ch] := 0;
	aWaiting[ch] := FALSE;
	aWaitAlarmId[ch] := 0;
	fbSetMacro[ch].Start := FALSE;
	fbWaitMacro[ch].Start := FALSE;

	IF aNciToPlc[ch].HskMFuncReq = 1 AND NOT fbGrantHold[ch].Q THEN
		bGrant := FALSE;
		nMFunc := TO_UINT(aNciToPlc[ch].HskMFuncNo);

		// Riga della tabella per (canale, M)
		nDef := -1;
		i := LOWER_BOUND(aDef, 1);
		WHILE i < LOWER_BOUND(aDef, 1) + nDefCount AND_THEN i <= UPPER_BOUND(aDef, 1) DO
			IF aDef[i].nChannel = ch AND aDef[i].nMFunc = nMFunc THEN
				nDef := i;
				EXIT;
			END_IF
			i := i + 1;
		END_WHILE

		IF nDef < 0 THEN
			// Senza riga il canale resterebbe fermo per sempre.
			IF bCycleRunning THEN
				aAlarmId[ch] := nUnknownAlarmId;
				aAlarmInfo[ch] := (ch + 1) * 1000 + nMFunc;
				bAbort := TRUE;
			END_IF
		ELSE
			stDef := aDef[nDef];

			CASE stDef.eKind OF
				E_MFuncKind.Nop:
					bGrant := TRUE;

				E_MFuncKind.LineNo:
					aLineNo[ch] := DINT_TO_UDINT(ItpGetHParam(aNciToPlc[ch]));
					bGrant := TRUE;

				E_MFuncKind.WaitStart:
					bGrant := bStart;

				E_MFuncKind.WaitH:
					fbWaitMacro[ch].Start := TRUE;
					fbWaitMacro[ch].WaitTime := DINT_TO_TIME(ItpGetHParam(aNciToPlc[ch]));
					IF fbWaitMacro[ch].Done THEN
						fbWaitMacro[ch].Start := FALSE;
						bGrant := TRUE;
					END_IF

				E_MFuncKind.Sync:
					dwSyncFlags := (dwSyncFlags OR stDef.dwSetWhileWaiting) AND NOT stDef.dwClearWhileWaiting;
					IF (dwSyncFlags AND stDef.dwWaitSet) = stDef.dwWaitSet AND (dwSyncFlags AND stDef.dwWaitClear) = 0 THEN
						dwSyncFlags := (dwSyncFlags OR stDef.dwSetOnGrant) AND NOT stDef.dwClearOnGrant;
						bGrant := TRUE;
					ELSE
						aWaiting[ch] := stDef.nWaitAlarmId <> 0;
						aWaitAlarmId[ch] := stDef.nWaitAlarmId;
					END_IF

				E_MFuncKind.ValveDirect:
					stValve := aValve[stDef.nValve];
					IF stDef.eAction = OUTPUT_ACTION_ENUM.SET THEN
						stValve.pSet^ := TRUE;
						IF stValve.eType = OUTPUT_ENUM.BISTABLE THEN
							stValve.pReset^ := FALSE;
						END_IF
					ELSE
						stValve.pSet^ := FALSE;
						IF stValve.eType = OUTPUT_ENUM.BISTABLE THEN
							stValve.pReset^ := TRUE;
						END_IF
					END_IF
					bGrant := TRUE;

				E_MFuncKind.Valve:
					IF stDef.nInterlock = 0 OR_ELSE aInterlock[stDef.nInterlock] THEN
						stValve := aValve[stDef.nValve];
						fbSetMacro[ch].Start := TRUE;
						fbSetMacro[ch].OutputType := stValve.eType;
						fbSetMacro[ch].ActionType := stDef.eAction;
						fbSetMacro[ch].TimeOutTime := stDef.tTimeout;
						IF stDef.bPostDelayFromH THEN
							fbSetMacro[ch].PostDelay := DINT_TO_TIME(ItpGetHParam(aNciToPlc[ch]));
						ELSE
							fbSetMacro[ch].PostDelay := stDef.tPostDelay;
						END_IF
						IF stDef.eAction = OUTPUT_ACTION_ENUM.SET THEN
							fbSetMacro[ch].FeedBack := stValve.pFbSet;
						ELSE
							fbSetMacro[ch].FeedBack := stValve.pFbReset;
						END_IF
						fbSetMacro[ch].SetOutput := stValve.pSet;
						IF stValve.pReset <> 0 THEN
							fbSetMacro[ch].ResetOutput := stValve.pReset;
						ELSE
							// SetMacro azzera ResetOutput^ anche per le monostabili quando va in timeout
							fbSetMacro[ch].ResetOutput := ADR(aNoResetOutput[ch]);
						END_IF

						IF fbSetMacro[ch].Done THEN
							fbSetMacro[ch].Start := FALSE;
							bGrant := TRUE;
						END_IF

						IF fbSetMacro[ch].Error THEN
							CASE stDef.eOnError OF
								E_MFuncOnError.Abort:
									aAlarmId[ch] := stDef.nAlarmId;
									aAlarmInfo[ch] := nMFunc;
									bAbort := TRUE;
								E_MFuncOnError.Grant:
									bGrant := TRUE;
							END_CASE
						END_IF
					ELSE
						aWaiting[ch] := stDef.nWaitAlarmId <> 0;
						aWaitAlarmId[ch] := stDef.nWaitAlarmId;
					END_IF
			END_CASE
		END_IF

		IF bGrant THEN
			aPlcToNci[ch].MFuncGranted := 1;
		END_IF
	ELSE
		aPlcToNci[ch].MFuncGranted := 0;
	END_IF
END_FOR

// Come prima in MAIN.AxisFunctionBlocks: le macro girano dopo la decisione, poi il fronte della
// concessione apre la finestra di 10 ms in cui il canale non viene servito.
FOR ch := 0 TO Core_Param.MAX_CHANNEL - 1 DO
	fbSetMacro[ch]();
	fbWaitMacro[ch]();
	fbGrantTrig[ch](CLK := aPlcToNci[ch].MFuncGranted = 1);
	fbGrantHold[ch](IN := fbGrantTrig[ch].Q, PT := T#10MS);
END_FOR

END_FUNCTION_BLOCK

// ---- Core/Valves/SetMacro.TcPOU
{attribute 'hide_all_locals'}
FUNCTION_BLOCK SetMacro
VAR_INPUT
	Start 							: BOOL;
	OutputType 						: OUTPUT_ENUM;
	ActionType						: OUTPUT_ACTION_ENUM;
	TimeOutTime						: TIME;
	PostDelay						: TIME;
	FeedBack						: POINTER TO BOOL;
	SetOutput 						: POINTER TO BOOL;
	ResetOutput 					: POINTER TO BOOL;
END_VAR

VAR_OUTPUT
	Busy 							: BOOL;
	Done							: BOOL;
	Error 							: BOOL;
END_VAR
VAR
	state 							: UINT;
	fbStartTrigger					: R_TRIG;
	startTriggerOutput				: BOOL;
	fbTimerOn 						: TON;
	fbTimerOnStart					: BOOL;
	fbTimerOnEnd 					: BOOL;
	fbPostTimer						: TON;
	fbPostTimerOnStart				: BOOL;
	fbPostTimerOnEnd				: BOOL;
END_VAR

fbTimerOn(IN:=fbTimerOnStart, PT := TimeOutTime, Q => fbTimerOnEnd);
fbPostTimer(IN:=fbPostTimerOnStart, PT := PostDelay, Q => fbPostTimerOnEnd);
fbStartTrigger(CLK := Start, Q => startTriggerOutput);

CASE state OF
	(************************** state 0 - IDLE *************************)  
	0:	
		Busy := FALSE;
		Done := FALSE;
		Error := FALSE;
		
		IF startTriggerOutput THEN
			Busy := TRUE;
			Error := FALSE;
			fbTimerOnStart := FALSE;
			state := 10;
		END_IF
	10:
		IF FeedBack^ THEN
			IF PostDelay <> T#0MS THEN
				fbPostTimerOnStart := TRUE;
				state := 30;
			ELSE
				state := 100;
			END_IF
		ELSE
			fbTimerOnStart := TRUE;
			state := 20;
		END_IF
	
	(************** state 20 - Set Output and wait for feedback *************)  
	20:
		CASE ActionType OF
			OUTPUT_ACTION_ENUM.SET:
				SetOutput^ := TRUE;
				IF OutputType = OUTPUT_ENUM.BISTABLE THEN
					ResetOutput^ := FALSE;
				END_IF

			OUTPUT_ACTION_ENUM.RESET:
				SetOutput^ := FALSE;
				IF OutputType = OUTPUT_ENUM.BISTABLE THEN
					ResetOutput^ := TRUE;
				END_IF
		END_CASE
		
		// Il timeout prevale anche se il feedback arriva nella stessa scansione.
		IF fbTimerOnEnd THEN
			fbTimerOnStart := FALSE;
			SetOutput^ := FALSE;
			ResetOutput^ := FALSE;
			state := 200;
		ELSIF FeedBack^ THEN
			fbTimerOnStart := FALSE;
			//SetOutput^ := FALSE;
			//ResetOutput^ := FALSE;
			
			IF PostDelay <> T#0MS THEN
				fbPostTimerOnStart := TRUE;
				state := 30;
			ELSE
				state := 100;
			END_IF
		END_IF
		
	(************** state 30 - Wait Post Time Delay *************)  
	30:
		IF fbPostTimerOnEnd THEN
			fbPostTimerOnStart := FALSE;
			state := 100;
		END_IF
	
	(************** state 100 - End *************)  
	100:
		Done := TRUE;
		state := 0;
	
	(************** state 100 - Error *************)  
	200:
		state := 0;
		Error := TRUE;
		
END_CASE

END_FUNCTION_BLOCK

// ---- Core/Valves/WaitMacro.TcPOU
FUNCTION_BLOCK WaitMacro
VAR_INPUT
	Start 							: BOOL;
	WaitTime						: TIME;
END_VAR
VAR_OUTPUT
	Busy 							: BOOL;
	Done							: BOOL;
END_VAR
VAR
	state 							: UINT;
	fbStartTrigger					: R_TRIG;
	startTriggerOutput				: BOOL;
	fbTimerOn 						: TON;
	fbTimerOnStart					: BOOL;
	fbTimerOnEnd 					: BOOL;
END_VAR

fbTimerOn(IN:=fbTimerOnStart, PT := WaitTime, Q => fbTimerOnEnd);
fbStartTrigger(CLK := Start, Q => startTriggerOutput);
		
CASE state OF
	(************************** state 0 - IDLE *************************)  
	0:	
		Busy := FALSE;
		Done := FALSE;
		
		IF startTriggerOutput THEN
			Busy := TRUE;
			fbTimerOnStart := TRUE;
			state := 10;
		END_IF
	10:
		IF fbTimerOnEnd OR (WaitTime = T#0MS) THEN
			fbTimerOnStart := FALSE;
			state := 100;
		END_IF
	
	(************** state 100 - End *************)  
	100:
		Done := TRUE;
		state := 0;
		
END_CASE

END_FUNCTION_BLOCK

// ---- Core/Diag/FB_DiagLog.TcPOU
// Storico dei cambi di passo del ciclo. Va chiamato una volta per ciclo PLC, dopo tutto cio' che puo'
// cambiare il passo (macchina a stati, funzioni M, allarmi), con stDiag.aChannel gia' aggiornato.
// Non conosce la macchina: riceve il passo, la sequenza e l'ultimo allarme come numeri.
FUNCTION_BLOCK FB_DiagLog
VAR_INPUT
	nState			: UINT;		// passo attuale del ciclo
	nSeqIdx			: UINT;		// sequenza corrente
	nAbortState		: UINT;		// passo che vale come abort: il suo evento si copia in stLastAbort
	nAlarmCount		: UDINT;	// quante volte e' stato memorizzato un allarme (cresce a ogni RaiseAlarm)
	nAlarmId		: UINT;		// ultimo allarme memorizzato
	nAlarmInfo		: UDINT;	// suo dettaglio
END_VAR
VAR_IN_OUT
	stDiag			: ST_Diag;	// aChannel, nSeqCount ed eCycleEndReason li scrive chi chiama
END_VAR
VAR
	bInit			: BOOL;
	tStateSince		: TIME;
	nAlarmCountSeen	: UDINT;
	stEvent			: ST_DiagEvent;
	i				: UINT;
END_VAR

IF NOT bInit THEN
	bInit := TRUE;
	stDiag.nState := nState;
	stDiag.nPrevState := nState;
	tStateSince := TIME();
	nAlarmCountSeen := nAlarmCount;
END_IF

IF nState <> stDiag.nState THEN
	stEvent.nIndex := stDiag.nEventCount + 1;
	stEvent.nTime := F_GetSystemTime();
	stEvent.nFromState := stDiag.nState;
	stEvent.nToState := nState;
	stEvent.nSeqIdx := nSeqIdx;

	FOR i := 0 TO Core_Param.MAX_CHANNEL - 1 DO
		stEvent.aLineNo[i] := stDiag.aChannel[i].nLineNo;
		IF stDiag.aChannel[i].bMWaiting THEN
			stEvent.aMFunc[i] := stDiag.aChannel[i].nMFunc;
		ELSE
			stEvent.aMFunc[i] := 0;
		END_IF
	END_FOR

	// Solo un allarme memorizzato dopo l'evento precedente: e' quello che ha causato questo cambio di passo.
	IF nAlarmCount <> nAlarmCountSeen THEN
		stEvent.nAlarmId := nAlarmId;
		stEvent.nAlarmInfo := nAlarmInfo;
		nAlarmCountSeen := nAlarmCount;
	ELSE
		stEvent.nAlarmId := 0;
		stEvent.nAlarmInfo := 0;
	END_IF

	stDiag.aEvent[stDiag.nEventCount MOD Core_Param.DIAG_EVENTS] := stEvent;
	stDiag.nEventCount := stDiag.nEventCount + 1;

	IF nState = nAbortState THEN
		stDiag.stLastAbort := stEvent;
	END_IF

	stDiag.nPrevState := stDiag.nState;
	stDiag.nState := nState;
	tStateSince := TIME();
END_IF

stDiag.tInState := TIME() - tStateSince;
stDiag.nSeqIdx := nSeqIdx;

END_FUNCTION_BLOCK

// ---- POUs/Clock.TcPOU
PROGRAM Clock
VAR
	{attribute 'hide'} 
	fbClock1OnHz 		: TON;
	{attribute 'hide'} 
	fbClock1OffHz 		: TON;
	{attribute 'hide'} 
	fbClock2OnHz 		: TON;
	{attribute 'hide'} 
	fbClock2OffHz 		: TON;
	{attribute 'hide'} 
	fbClock5OnHz 		: TON;
	{attribute 'hide'} 
	fbClock5OffHz 		: TON;
	{attribute 'hide'} 
	etClockOn2Hz		: TIME;
	{attribute 'hide'} 
	etClockOff2Hz		: TIME;
	{attribute 'hide'} 
	etClockOn1Hz		: TIME;
	{attribute 'hide'} 
	etClockOff1Hz		: TIME;
	{attribute 'hide'} 
	etClockOn5Hz		: TIME;
	{attribute 'hide'} 
	etClockOff5Hz		: TIME;
	pulse1Hz			: BOOL;
	pulse2Hz			: BOOL;
	pulse5Hz			: BOOL;
	{attribute 'hide'} 
	fbClockSr1Hz		: SR;
	{attribute 'hide'} 
	fbClockSr2Hz		: SR;
	{attribute 'hide'} 
	fbClockSr5Hz		: SR;
END_VAR

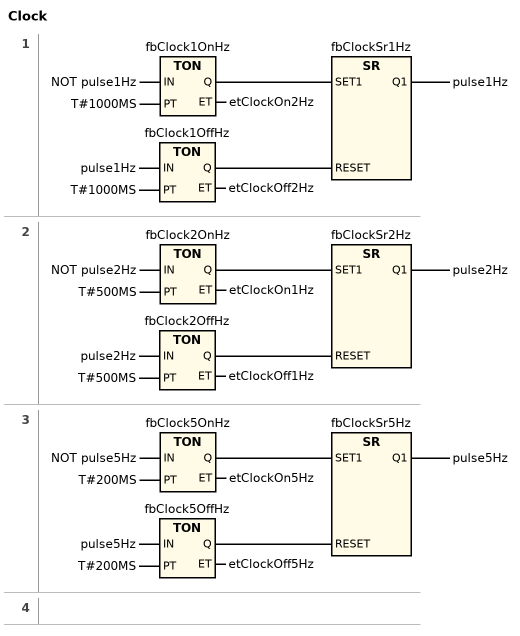
// NETWORK 1
fbClock1OnHz(IN := NOT pulse1Hz, PT := T#1000MS, ET => etClockOn2Hz); // TON
fbClock1OffHz(IN := pulse1Hz, PT := T#1000MS, ET => etClockOff2Hz); // TON
fbClockSr1Hz(SET1 := fbClock1OnHz.Q, RESET := fbClock1OffHz.Q); // SR
pulse1Hz := fbClockSr1Hz.Q1;

// NETWORK 2
fbClock2OnHz(IN := NOT pulse2Hz, PT := T#500MS, ET => etClockOn1Hz); // TON
fbClock2OffHz(IN := pulse2Hz, PT := T#500MS, ET => etClockOff1Hz); // TON
fbClockSr2Hz(SET1 := fbClock2OnHz.Q, RESET := fbClock2OffHz.Q); // SR
pulse2Hz := fbClockSr2Hz.Q1;

// NETWORK 3
fbClock5OnHz(IN := NOT pulse5Hz, PT := T#200MS, ET => etClockOn5Hz); // TON
fbClock5OffHz(IN := pulse5Hz, PT := T#200MS, ET => etClockOff5Hz); // TON
fbClockSr5Hz(SET1 := fbClock5OnHz.Q, RESET := fbClock5OffHz.Q); // SR
pulse5Hz := fbClockSr5Hz.Q1;

// NETWORK 4

END_PROGRAM

// ---- POUs/Messages/ClearAlarms.TcPOU
// Reset: azzera tutti gli allarmi. Quelli a livello ancora presenti vengono riattivati
// da MAIN.AlarmManager nello stesso ciclo (e' chiamata dopo la macchina a stati).
FUNCTION ClearAlarms : BOOL

MEMSET(ADR(Alarms.Active), 0, SIZEOF(Alarms.Active));
MEMSET(ADR(Alarms.Info), 0, SIZEOF(Alarms.Info));
ClearAlarms := TRUE;

END_FUNCTION
